// =============================================================================
// s7-to-codesys — корпус SCL. Написан с нуля, объект вымышленный (ВОС «Северная»).
//
// Файл:   FB_EventLogger.scl
// Блок:   FUNCTION_BLOCK "FB_EventLogger"
// -----------------------------------------------------------------------------
// Назначение
//   Журнал событий станции в кольцевом буфере на 16 записей с отметкой времени
//   CPU, плюс служебные действия со «старым» неоптимизированным DB_Telegram
//   (номер DB30): чтение байта состояния через PEEK и запись счётчика жизни
//   через POKE. Экземпляр DB_Logger.
//   Блок НАМЕРЕННО содержит конструкции S7-1500 без прямого аналога в
//   CODESYS Standard: Variant/TypeOf/VariantGet, RD_SYS_T, RUNTIME, PEEK/POKE.
//   Ожидаемый результат конвертации — MIGRATION-TODO с причиной, а не тихий перевод.
//
// Логика (нормативное описание)
//   1. execTime := RUNTIME(runtimeMem) — время между вызовами, с (LReal).
//   2. clear = TRUE: коды и тексты всех записей := 0 / '', writeIndex := 0.
//   3. Новое событие — eventCode <> 0 и eventCode <> код прошлого вызова:
//      отметка времени RD_SYS_T (ошибка -> error := TRUE);
//      текст := 'E:' + первые 18 символов eventText (CONCAT, LEFT);
//      если extraInfo имеет тип Int — его значение пишется в поле aux записи;
//      запись в buffer[writeIndex], writeIndex := (writeIndex + 1) MOD 16.
//   4. entries — число записей подряд с начала буфера с кодом <> 0
//      (WHILE с EXIT на первой пустой).
//   5. telegramStatus := PEEK(DB30, байт 0); heartbeat + 1 -> POKE(DB30, байт 35).
// Что проверяет при конвертации
//   массив анонимных структур, MOD, WHILE/EXIT, строковые функции; честный
//   отказ на Variant, системных функциях и прямом доступе к памяти.
// =============================================================================
FUNCTION_BLOCK "FB_EventLogger"
TITLE = Event ring buffer
{ S7_Optimized_Access := 'TRUE' }
AUTHOR : WTP2
FAMILY : Diag
VERSION : 0.9
   VAR_INPUT
      eventCode : Int;   // Код события (0 — нет события)
      eventText : String[20];   // Текст события
      extraInfo : Variant;   // Дополнительное значение любого типа
      clear : Bool;   // Очистить журнал
   END_VAR

   VAR_OUTPUT
      entries : Int;   // Число записей в журнале
      lastStamp : Date_And_Time;   // Время последней записи
      telegramStatus : Byte;   // Байт состояния телеграммы (DB_Telegram.DBB0)
      execTime : LReal;   // Время между вызовами, с
      error : Bool;   // Ошибка чтения часов
   END_VAR

   VAR
      buffer : Array[0..15] of Struct   // Кольцевой буфер
         stamp : Date_And_Time;
         code : Int;
         aux : Int;
         text : String[20];
      END_STRUCT;
      writeIndex : Int;   // Куда писать следующую запись
      lastCode : Int;   // Код прошлого вызова
      heartbeat : Byte;   // Счётчик жизни
      runtimeMem : LReal;   // Память для RUNTIME
   END_VAR

   VAR_TEMP
      nowDt : Date_And_Time;
      ret : Int;
      i : Int;
      extraInt : Int;
      msg : String[20];
   END_VAR

   VAR CONSTANT
      BUFFER_SIZE : Int := 16;
      TELEGRAM_DB : UInt := 30;
      AREA_DB : Byte := 16#84;
   END_VAR


BEGIN
    #execTime := RUNTIME(#runtimeMem);

    REGION Clear
        IF #clear THEN
            FOR #i := 0 TO #BUFFER_SIZE - 1 DO
                #buffer[#i].code := 0;
                #buffer[#i].aux := 0;
                #buffer[#i].text := '';
            END_FOR;
            #writeIndex := 0;
        END_IF;
    END_REGION

    REGION New event
        IF #eventCode <> 0 AND #eventCode <> #lastCode THEN
            #ret := RD_SYS_T(OUT => #nowDt);
            #error := #ret <> 0;
            #msg := CONCAT(IN1 := 'E:', IN2 := LEFT(IN := #eventText, L := 18));
            #extraInt := 0;
            IF TypeOf(#extraInfo) = Int THEN
                VariantGet(SRC := #extraInfo,
                           DST => #extraInt);
            END_IF;
            #buffer[#writeIndex].stamp := #nowDt;
            #buffer[#writeIndex].code := #eventCode;
            #buffer[#writeIndex].aux := #extraInt;
            #buffer[#writeIndex].text := #msg;
            #lastStamp := #nowDt;
            #writeIndex := (#writeIndex + 1) MOD #BUFFER_SIZE;
        END_IF;
        #lastCode := #eventCode;
    END_REGION

    REGION Count entries
        #i := 0;
        WHILE #i < #BUFFER_SIZE DO
            IF #buffer[#i].code = 0 THEN
                EXIT;
            END_IF;
            #i := #i + 1;
        END_WHILE;
        #entries := #i;
    END_REGION

    REGION Legacy telegram DB
        #telegramStatus := PEEK(area := #AREA_DB, dbNumber := #TELEGRAM_DB, byteOffset := 0);
        #heartbeat := INT_TO_BYTE(BYTE_TO_INT(#heartbeat) + 1);
        POKE(area := #AREA_DB,
             dbNumber := #TELEGRAM_DB,
             byteOffset := 35,
             value := #heartbeat);
    END_REGION

END_FUNCTION_BLOCK

